Fanuc KAREL source: kb00033.KL

PROGRAM KB00033
%STACKSIZE=65535
%PRIORITY=65535
%NOLOCKGROUP
VAR
P2 : STRING[80]
P3 : INTEGER
-- UNRESOLVED DECLARATIONS (source type spelling not recovered)
-- P1 : TYPE_0x001C (type_u16=0x001C)
BEGIN
P2='A'
P3=1
CNV_CNF_STRG(P1,P2,P3,1)
END KB00033
